// CFC twin of T_SafeDecouple_Tests: the same tests drawn as CFC diagrams, the way a TwinSAFE project is authored.
    FUNCTION_BLOCK T_SafeDecouple_Tests_CFC EXTENDS T_SafeCfcTestSuite
    VAR
    // Test_InputsLoopedToOutputsOnlyWhenRunning
    group_1 : T_SafeGroup;
    fb_1 : T_SafeDecouple(group := group_1);
END_VAR

Test_InputsLoopedToOutputsOnlyWhenRunning();

METHOD PRIVATE Test_InputsLoopedToOutputsOnlyWhenRunning
// note: this text did not pass the execution check against the stored diagram
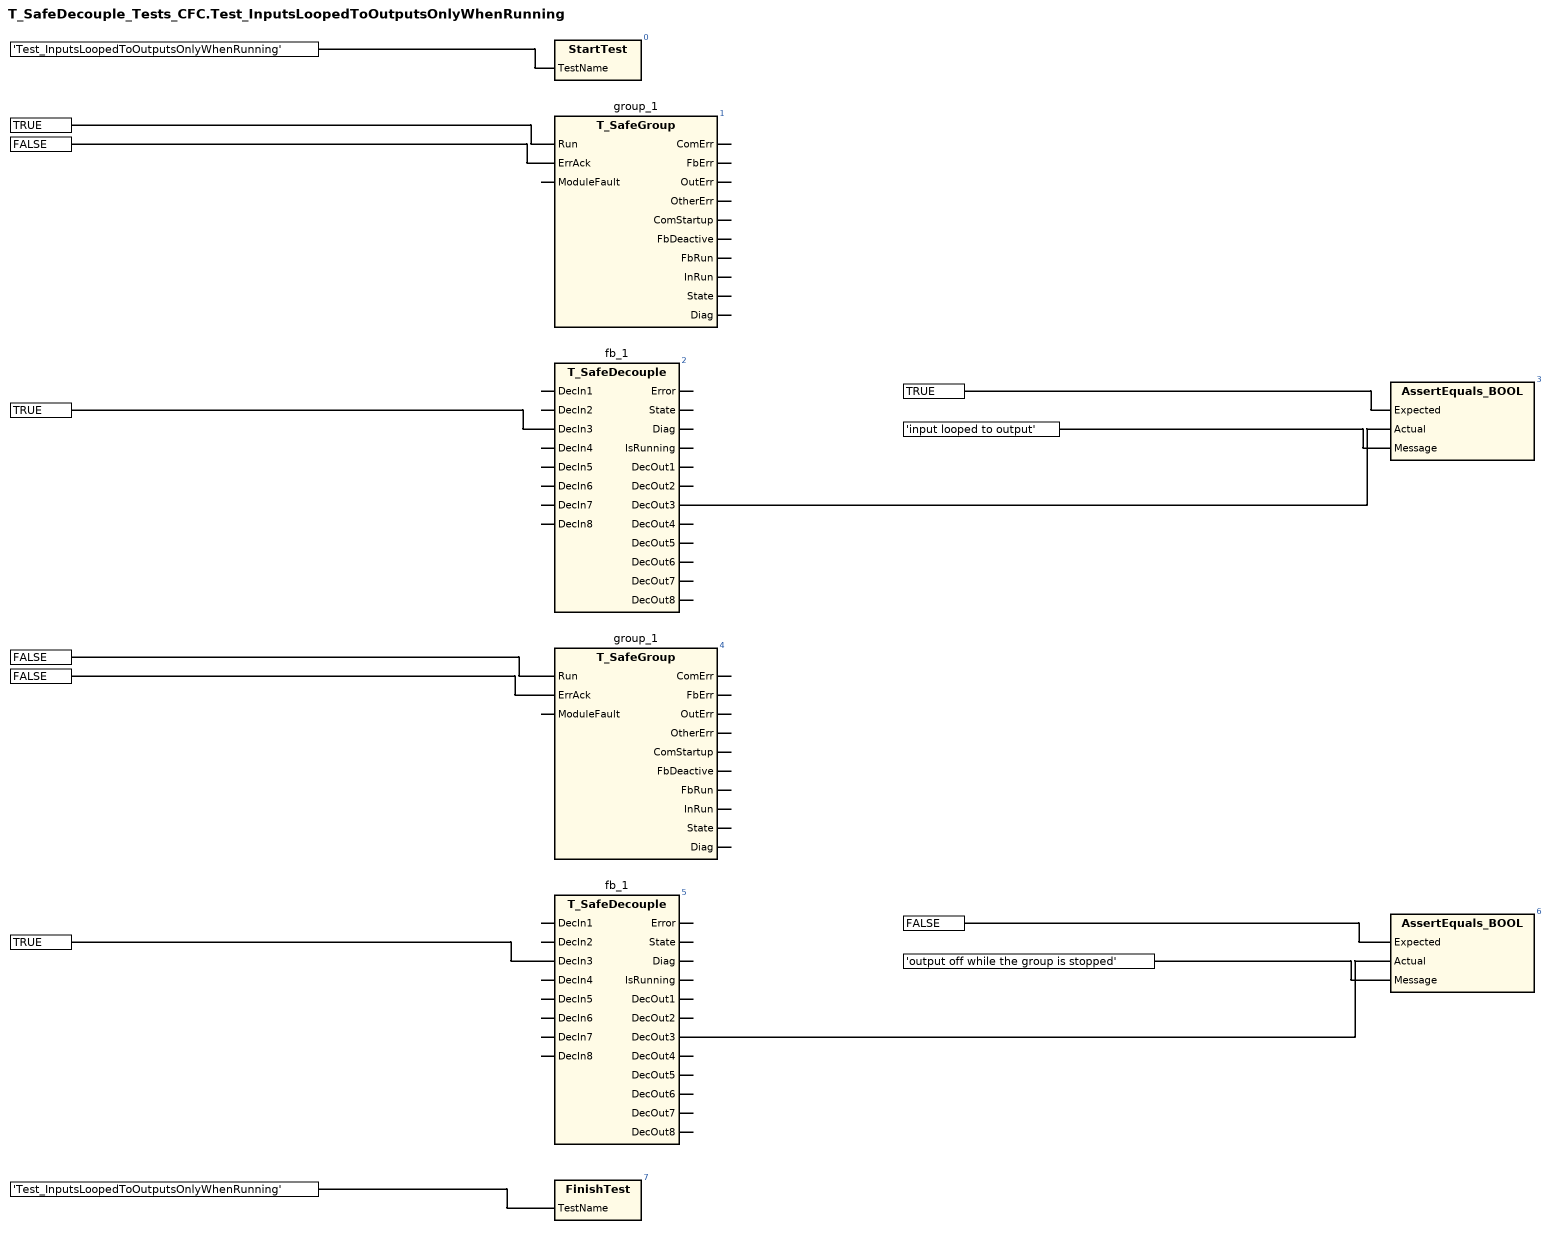
StartTest(TestName := 'Test_InputsLoopedToOutputsOnlyWhenRunning');
group_1(Run := TRUE, ErrAck := FALSE); // T_SafeGroup
fb_1(DecIn3 := TRUE); // T_SafeDecouple
AssertEquals_BOOL(Expected := TRUE, Actual := fb_1.DecOut3, Message := 'input looped to output');
group_1(Run := FALSE, ErrAck := FALSE); // T_SafeGroup
fb_1(DecIn3 := TRUE); // T_SafeDecouple
AssertEquals_BOOL(Expected := FALSE, Actual := fb_1.DecOut3, Message := 'output off while the group is stopped');
FinishTest(TestName := 'Test_InputsLoopedToOutputsOnlyWhenRunning');
END_METHOD

END_FUNCTION_BLOCK

(* stored: Version 1.1.0.1, ProductVersion 3.1.4026.22
   POU T_SafeDecouple_Tests_CFC: Id {901187d0-da6d-5001-b298-1307acc58f68}, SpecialFunc None
   Method Test_InputsLoopedToOutputsOnlyWhenRunning: Id {bd4e4555-f336-5510-8a6e-cbbb007d6548} *)
